Fanuc KAREL source: kb00044.KL

-- PROVISIONAL review KL for V940-1; original PC SHA256 463385d52d9acd5178af6be934f223b7615a28d1c3df33b263db40f5b198cdcf
-- Incomplete behavior may be omitted. Consult companion uncertainty JSON. Do not deploy.
PROGRAM KB00044
%NOLOCKGROUP
BEGIN
  -- V9_ZERO_TABLE_METADATA_HINT layout=0002_ascii; no indexed target words; source/name/runtime held
  -- UNRESOLVED_PC offsets 5-14; opcodes 3F,75
  -- UNRESOLVED_PC offsets 19-28; opcodes 3F,75
  -- UNRESOLVED_PC offsets 33-40; opcodes 9D,23
  -- UNRESOLVED_PC offsets 45-52; opcodes 9D,23
  -- UNRESOLVED_PC offsets 57-64; opcodes 9D,23
  -- UNRESOLVED_PC offsets 69-113; opcodes 27,22,2A,22,2A,22,22,22,22,31
  -- UNRESOLVED_PC offsets 118-122; opcodes 7F
END KB00044
